Fanuc KAREL source: kt00293.KL

-- PROVISIONAL review KL for V770-1; original PC SHA256 d04c193cbe47158a5e5133aed8266c33d50cdc1ad707cca72c5b784635ce8e2f
-- Incomplete behavior may be omitted. Consult companion uncertainty JSON. Do not deploy.
PROGRAM KT00293
%NOLOCKGROUP
VAR
  I1 : INTEGER
  I2 : INTEGER
  OUT : BOOLEAN
BEGIN
  -- UNRESOLVED_PC offsets 5-16; opcodes 2E,23
  -- UNRESOLVED_PC offsets 21-32; opcodes 2E,23
  -- UNRESOLVED_PC offsets 37-48; opcodes 2E,23
  -- UNRESOLVED_PC offsets 53-64; opcodes 2E,23
  -- UNRESOLVED_PC offsets 69-88; opcodes 21,21,58,23
  -- UNRESOLVED_PC offsets 93-97; opcodes 7F
END KT00293
